// TIA Portal V20 export
Screen "170PRBCompleteDisplay"  1276x673
  ScreenItem "sequenceControlFaceplate_Lite_1" at 380,555 size 641x64  Type=HmiFaceplateContainer
  ScreenItem "Title_ScreenOverview_X390_Y2" at 390,2 size 500x30  Type=HmiTextBox
  ScreenItem "Button_Back_1" at 2,2 size 90x60  Type=HmiButton
  ScreenItem "Tec-Unit_LegendᆉY2" at 1183,2 size 90x60  Type=HmiButton
  ScreenItem "permanentareaborderrectangle" at 0,0 size 0x0  Type=HmiRectangle
  ScreenItem "面板容器_2" at 1091,4 size 88x58  Type=HmiFaceplateContainer
  ScreenItem "OPMode1_Blocked" at 1165,6 size 14x14  Type=HmiGraphicView
  ScreenItem "OPMode3_Foreground_Blocked" at 1090,5 size 88x58  Type=HmiGraphicView
  ScreenItem "Button_Back" at 2,4 size 90x60  Type=HmiButton
  ScreenItem "Title_ScreenOverview_X390_Y2_1" at 380,5 size 510x57  Type=HmiTextBox
  ScreenItem "面板容器_3" at 217,276 size 163x70  Type=HmiFaceplateContainer
  ScreenItem "面板容器_4" at 12,276 size 163x70  Type=HmiFaceplateContainer
